FUNCTION "FRK_PersistDirty" : Void
{ S7_Optimized_Access := 'TRUE' }
VERSION : 0.1
VAR_INPUT
    Slot : Int;
END_VAR
VAR_TEMP
    Stamp : LDT;
    NativeResult : Int;
END_VAR
BEGIN
    IF #Slot < 1 OR #Slot > 20 THEN RETURN; END_IF;
    IF NOT "FRK_PersistConsumers".Rows[#Slot].Dirty THEN
        #NativeResult := RD_SYS_T(OUT => #Stamp);
        IF "FRK_PersistConsumers".Rows[#Slot].Ticket = 0 THEN "FRK_PersistConsumers".Rows[#Slot].PendingSince := #Stamp;
        ELSE "FRK_PersistConsumers".Rows[#Slot].NextSince := #Stamp; END_IF;
    END_IF;
    "FRK_PersistConsumers".Rows[#Slot].Dirty := TRUE;
END_FUNCTION
FUNCTION "FRK_PersistConfigSlot" : Int
{ S7_Optimized_Access := 'TRUE' }
VERSION : 0.1
VAR_INPUT
    Scope : String;
    ModelCode : String;
    Kind : DInt;
END_VAR
BEGIN
    #FRK_PersistConfigSlot := 0;
    IF #Scope = 'StationA' AND #ModelCode = '' AND #Kind = 1 THEN #FRK_PersistConfigSlot := 1; RETURN; END_IF;
    IF #Scope = 'StationA' AND #ModelCode = '' AND #Kind = 1 THEN #FRK_PersistConfigSlot := 1; RETURN; END_IF;
    IF #Scope = 'StationA' AND #ModelCode = '' AND #Kind = 1 THEN #FRK_PersistConfigSlot := 1; RETURN; END_IF;
    IF #Scope = 'StationA' AND #ModelCode = '' AND #Kind = 1 THEN #FRK_PersistConfigSlot := 1; RETURN; END_IF;
    IF #Scope = 'StationA' AND #ModelCode = '' AND #Kind = 1 THEN #FRK_PersistConfigSlot := 1; RETURN; END_IF;
    IF #Scope = 'StationA' AND #ModelCode = '' AND #Kind = 1 THEN #FRK_PersistConfigSlot := 1; RETURN; END_IF;
    IF #Scope = 'StationA' AND #ModelCode = '' AND #Kind = 1 THEN #FRK_PersistConfigSlot := 1; RETURN; END_IF;
    IF #Scope = 'StationA' AND #ModelCode = '' AND #Kind = 1 THEN #FRK_PersistConfigSlot := 1; RETURN; END_IF;
    IF #Scope = 'StationA.Satellite' AND #ModelCode = '' AND #Kind = 1 THEN #FRK_PersistConfigSlot := 1; RETURN; END_IF;
    IF #Scope = 'StationA.Satellite' AND #ModelCode = '' AND #Kind = 1 THEN #FRK_PersistConfigSlot := 1; RETURN; END_IF;
    IF #Scope = 'StationA.Satellite' AND #ModelCode = '' AND #Kind = 1 THEN #FRK_PersistConfigSlot := 1; RETURN; END_IF;
    IF #Scope = 'StationA.Satellite' AND #ModelCode = '' AND #Kind = 1 THEN #FRK_PersistConfigSlot := 1; RETURN; END_IF;
    IF #Scope = 'StationA.Satellite' AND #ModelCode = '' AND #Kind = 1 THEN #FRK_PersistConfigSlot := 1; RETURN; END_IF;
    IF #Scope = 'StationA.Satellite' AND #ModelCode = '' AND #Kind = 1 THEN #FRK_PersistConfigSlot := 1; RETURN; END_IF;
    IF #Scope = 'StationA.Satellite' AND #ModelCode = '' AND #Kind = 1 THEN #FRK_PersistConfigSlot := 1; RETURN; END_IF;
    IF #Scope = 'StationA.Satellite' AND #ModelCode = '' AND #Kind = 1 THEN #FRK_PersistConfigSlot := 1; RETURN; END_IF;
    IF #Scope = 'StationA.Satellite' AND #ModelCode = '' AND #Kind = 1 THEN #FRK_PersistConfigSlot := 1; RETURN; END_IF;
    IF #Scope = 'StationA.Satellite' AND #ModelCode = '' AND #Kind = 1 THEN #FRK_PersistConfigSlot := 1; RETURN; END_IF;
    IF #Scope = 'StationA.Satellite.Inner' AND #ModelCode = '' AND #Kind = 1 THEN #FRK_PersistConfigSlot := 1; RETURN; END_IF;
    IF #Scope = 'StationA.Satellite.Inner' AND #ModelCode = '' AND #Kind = 1 THEN #FRK_PersistConfigSlot := 1; RETURN; END_IF;
    IF #Scope = 'StationA.Satellite.Inner' AND #ModelCode = '' AND #Kind = 1 THEN #FRK_PersistConfigSlot := 1; RETURN; END_IF;
    IF #Scope = 'StationA.Satellite.Inner' AND #ModelCode = '' AND #Kind = 1 THEN #FRK_PersistConfigSlot := 1; RETURN; END_IF;
    IF #Scope = 'StationA.Satellite.Inner' AND #ModelCode = '' AND #Kind = 1 THEN #FRK_PersistConfigSlot := 1; RETURN; END_IF;
    IF #Scope = 'StationA.Satellite.Inner' AND #ModelCode = '' AND #Kind = 1 THEN #FRK_PersistConfigSlot := 1; RETURN; END_IF;
    IF #Scope = 'StationA.Satellite.Inner' AND #ModelCode = '' AND #Kind = 1 THEN #FRK_PersistConfigSlot := 1; RETURN; END_IF;
    IF #Scope = 'StationA.Satellite.Inner' AND #ModelCode = '' AND #Kind = 1 THEN #FRK_PersistConfigSlot := 1; RETURN; END_IF;
    IF #Scope = 'StationA.Satellite.Inner' AND #ModelCode = '' AND #Kind = 1 THEN #FRK_PersistConfigSlot := 1; RETURN; END_IF;
    IF #Scope = 'StationA.Satellite.Inner' AND #ModelCode = '' AND #Kind = 1 THEN #FRK_PersistConfigSlot := 1; RETURN; END_IF;
    IF #Scope = 'StationA' AND #ModelCode = 'MODEL_A' AND #Kind = 0 THEN #FRK_PersistConfigSlot := 2; RETURN; END_IF;
    IF #Scope = 'StationA' AND #ModelCode = 'MODEL_A' AND #Kind = 0 THEN #FRK_PersistConfigSlot := 2; RETURN; END_IF;
    IF #Scope = 'StationA' AND #ModelCode = 'MODEL_A' AND #Kind = 0 THEN #FRK_PersistConfigSlot := 2; RETURN; END_IF;
    IF #Scope = 'StationA' AND #ModelCode = 'MODEL_A' AND #Kind = 0 THEN #FRK_PersistConfigSlot := 2; RETURN; END_IF;
    IF #Scope = 'StationA.Cell' AND #ModelCode = 'MODEL_A' AND #Kind = 0 THEN #FRK_PersistConfigSlot := 2; RETURN; END_IF;
    IF #Scope = 'StationA.Cell' AND #ModelCode = 'MODEL_A' AND #Kind = 0 THEN #FRK_PersistConfigSlot := 2; RETURN; END_IF;
    IF #Scope = 'StationA.Cell.Clamp' AND #ModelCode = 'MODEL_A' AND #Kind = 0 THEN #FRK_PersistConfigSlot := 2; RETURN; END_IF;
    IF #Scope = 'StationA.Cell.Clamp' AND #ModelCode = 'MODEL_A' AND #Kind = 0 THEN #FRK_PersistConfigSlot := 2; RETURN; END_IF;
    IF #Scope = 'StationA.Cell.Gate' AND #ModelCode = 'MODEL_A' AND #Kind = 0 THEN #FRK_PersistConfigSlot := 2; RETURN; END_IF;
    IF #Scope = 'StationA.Cell.Gate' AND #ModelCode = 'MODEL_A' AND #Kind = 0 THEN #FRK_PersistConfigSlot := 2; RETURN; END_IF;
    IF #Scope = 'StationA.Satellite' AND #ModelCode = 'MODEL_A' AND #Kind = 0 THEN #FRK_PersistConfigSlot := 2; RETURN; END_IF;
    IF #Scope = 'StationA.Satellite' AND #ModelCode = 'MODEL_A' AND #Kind = 0 THEN #FRK_PersistConfigSlot := 2; RETURN; END_IF;
    IF #Scope = 'StationA.Satellite.Cell' AND #ModelCode = 'MODEL_A' AND #Kind = 0 THEN #FRK_PersistConfigSlot := 2; RETURN; END_IF;
    IF #Scope = 'StationA.Satellite.Cell' AND #ModelCode = 'MODEL_A' AND #Kind = 0 THEN #FRK_PersistConfigSlot := 2; RETURN; END_IF;
    IF #Scope = 'StationA.Satellite.Cell.Clamp' AND #ModelCode = 'MODEL_A' AND #Kind = 0 THEN #FRK_PersistConfigSlot := 2; RETURN; END_IF;
    IF #Scope = 'StationA.Satellite.Cell.Clamp' AND #ModelCode = 'MODEL_A' AND #Kind = 0 THEN #FRK_PersistConfigSlot := 2; RETURN; END_IF;
    IF #Scope = 'StationA.Satellite.Cell.Gate' AND #ModelCode = 'MODEL_A' AND #Kind = 0 THEN #FRK_PersistConfigSlot := 2; RETURN; END_IF;
    IF #Scope = 'StationA.Satellite.Cell.Gate' AND #ModelCode = 'MODEL_A' AND #Kind = 0 THEN #FRK_PersistConfigSlot := 2; RETURN; END_IF;
    IF #Scope = 'StationA.Satellite.Inner' AND #ModelCode = 'MODEL_A' AND #Kind = 0 THEN #FRK_PersistConfigSlot := 2; RETURN; END_IF;
    IF #Scope = 'StationA.Satellite.Inner' AND #ModelCode = 'MODEL_A' AND #Kind = 0 THEN #FRK_PersistConfigSlot := 2; RETURN; END_IF;
    IF #Scope = 'StationA.Satellite.Inner.Cell' AND #ModelCode = 'MODEL_A' AND #Kind = 0 THEN #FRK_PersistConfigSlot := 2; RETURN; END_IF;
    IF #Scope = 'StationA.Satellite.Inner.Cell' AND #ModelCode = 'MODEL_A' AND #Kind = 0 THEN #FRK_PersistConfigSlot := 2; RETURN; END_IF;
    IF #Scope = 'StationA.Satellite.Inner.Cell.Clamp' AND #ModelCode = 'MODEL_A' AND #Kind = 0 THEN #FRK_PersistConfigSlot := 2; RETURN; END_IF;
    IF #Scope = 'StationA.Satellite.Inner.Cell.Clamp' AND #ModelCode = 'MODEL_A' AND #Kind = 0 THEN #FRK_PersistConfigSlot := 2; RETURN; END_IF;
    IF #Scope = 'StationA.Satellite.Inner.Cell.Gate' AND #ModelCode = 'MODEL_A' AND #Kind = 0 THEN #FRK_PersistConfigSlot := 2; RETURN; END_IF;
    IF #Scope = 'StationA.Satellite.Inner.Cell.Gate' AND #ModelCode = 'MODEL_A' AND #Kind = 0 THEN #FRK_PersistConfigSlot := 2; RETURN; END_IF;
    IF #Scope = 'StationA' AND #ModelCode = 'MODEL_B' AND #Kind = 0 THEN #FRK_PersistConfigSlot := 3; RETURN; END_IF;
    IF #Scope = 'StationA' AND #ModelCode = 'MODEL_B' AND #Kind = 0 THEN #FRK_PersistConfigSlot := 3; RETURN; END_IF;
    IF #Scope = 'StationA' AND #ModelCode = 'MODEL_B' AND #Kind = 0 THEN #FRK_PersistConfigSlot := 3; RETURN; END_IF;
    IF #Scope = 'StationA' AND #ModelCode = 'MODEL_B' AND #Kind = 0 THEN #FRK_PersistConfigSlot := 3; RETURN; END_IF;
    IF #Scope = 'StationA.Cell' AND #ModelCode = 'MODEL_B' AND #Kind = 0 THEN #FRK_PersistConfigSlot := 3; RETURN; END_IF;
    IF #Scope = 'StationA.Cell' AND #ModelCode = 'MODEL_B' AND #Kind = 0 THEN #FRK_PersistConfigSlot := 3; RETURN; END_IF;
    IF #Scope = 'StationA.Cell.Clamp' AND #ModelCode = 'MODEL_B' AND #Kind = 0 THEN #FRK_PersistConfigSlot := 3; RETURN; END_IF;
    IF #Scope = 'StationA.Cell.Clamp' AND #ModelCode = 'MODEL_B' AND #Kind = 0 THEN #FRK_PersistConfigSlot := 3; RETURN; END_IF;
    IF #Scope = 'StationA.Cell.Gate' AND #ModelCode = 'MODEL_B' AND #Kind = 0 THEN #FRK_PersistConfigSlot := 3; RETURN; END_IF;
    IF #Scope = 'StationA.Cell.Gate' AND #ModelCode = 'MODEL_B' AND #Kind = 0 THEN #FRK_PersistConfigSlot := 3; RETURN; END_IF;
    IF #Scope = 'StationA.Satellite' AND #ModelCode = 'MODEL_B' AND #Kind = 0 THEN #FRK_PersistConfigSlot := 3; RETURN; END_IF;
    IF #Scope = 'StationA.Satellite' AND #ModelCode = 'MODEL_B' AND #Kind = 0 THEN #FRK_PersistConfigSlot := 3; RETURN; END_IF;
    IF #Scope = 'StationA.Satellite.Cell' AND #ModelCode = 'MODEL_B' AND #Kind = 0 THEN #FRK_PersistConfigSlot := 3; RETURN; END_IF;
    IF #Scope = 'StationA.Satellite.Cell' AND #ModelCode = 'MODEL_B' AND #Kind = 0 THEN #FRK_PersistConfigSlot := 3; RETURN; END_IF;
    IF #Scope = 'StationA.Satellite.Cell.Clamp' AND #ModelCode = 'MODEL_B' AND #Kind = 0 THEN #FRK_PersistConfigSlot := 3; RETURN; END_IF;
    IF #Scope = 'StationA.Satellite.Cell.Clamp' AND #ModelCode = 'MODEL_B' AND #Kind = 0 THEN #FRK_PersistConfigSlot := 3; RETURN; END_IF;
    IF #Scope = 'StationA.Satellite.Cell.Gate' AND #ModelCode = 'MODEL_B' AND #Kind = 0 THEN #FRK_PersistConfigSlot := 3; RETURN; END_IF;
    IF #Scope = 'StationA.Satellite.Cell.Gate' AND #ModelCode = 'MODEL_B' AND #Kind = 0 THEN #FRK_PersistConfigSlot := 3; RETURN; END_IF;
    IF #Scope = 'StationA.Satellite.Inner' AND #ModelCode = 'MODEL_B' AND #Kind = 0 THEN #FRK_PersistConfigSlot := 3; RETURN; END_IF;
    IF #Scope = 'StationA.Satellite.Inner' AND #ModelCode = 'MODEL_B' AND #Kind = 0 THEN #FRK_PersistConfigSlot := 3; RETURN; END_IF;
    IF #Scope = 'StationA.Satellite.Inner.Cell' AND #ModelCode = 'MODEL_B' AND #Kind = 0 THEN #FRK_PersistConfigSlot := 3; RETURN; END_IF;
    IF #Scope = 'StationA.Satellite.Inner.Cell' AND #ModelCode = 'MODEL_B' AND #Kind = 0 THEN #FRK_PersistConfigSlot := 3; RETURN; END_IF;
    IF #Scope = 'StationA.Satellite.Inner.Cell.Clamp' AND #ModelCode = 'MODEL_B' AND #Kind = 0 THEN #FRK_PersistConfigSlot := 3; RETURN; END_IF;
    IF #Scope = 'StationA.Satellite.Inner.Cell.Clamp' AND #ModelCode = 'MODEL_B' AND #Kind = 0 THEN #FRK_PersistConfigSlot := 3; RETURN; END_IF;
    IF #Scope = 'StationA.Satellite.Inner.Cell.Gate' AND #ModelCode = 'MODEL_B' AND #Kind = 0 THEN #FRK_PersistConfigSlot := 3; RETURN; END_IF;
    IF #Scope = 'StationA.Satellite.Inner.Cell.Gate' AND #ModelCode = 'MODEL_B' AND #Kind = 0 THEN #FRK_PersistConfigSlot := 3; RETURN; END_IF;
    IF #Scope = 'StationB' AND #ModelCode = '' AND #Kind = 1 THEN #FRK_PersistConfigSlot := 9; RETURN; END_IF;
    IF #Scope = 'StationB' AND #ModelCode = '' AND #Kind = 1 THEN #FRK_PersistConfigSlot := 9; RETURN; END_IF;
    IF #Scope = 'StationB' AND #ModelCode = '' AND #Kind = 1 THEN #FRK_PersistConfigSlot := 9; RETURN; END_IF;
    IF #Scope = 'StationB' AND #ModelCode = '' AND #Kind = 1 THEN #FRK_PersistConfigSlot := 9; RETURN; END_IF;
    IF #Scope = 'StationB' AND #ModelCode = '' AND #Kind = 1 THEN #FRK_PersistConfigSlot := 9; RETURN; END_IF;
    IF #Scope = 'StationB' AND #ModelCode = '' AND #Kind = 1 THEN #FRK_PersistConfigSlot := 9; RETURN; END_IF;
    IF #Scope = 'StationB' AND #ModelCode = '' AND #Kind = 1 THEN #FRK_PersistConfigSlot := 9; RETURN; END_IF;
    IF #Scope = 'StationB' AND #ModelCode = '' AND #Kind = 1 THEN #FRK_PersistConfigSlot := 9; RETURN; END_IF;
    IF #Scope = 'StationB.Satellite' AND #ModelCode = '' AND #Kind = 1 THEN #FRK_PersistConfigSlot := 9; RETURN; END_IF;
    IF #Scope = 'StationB.Satellite' AND #ModelCode = '' AND #Kind = 1 THEN #FRK_PersistConfigSlot := 9; RETURN; END_IF;
    IF #Scope = 'StationB.Satellite' AND #ModelCode = '' AND #Kind = 1 THEN #FRK_PersistConfigSlot := 9; RETURN; END_IF;
    IF #Scope = 'StationB.Satellite' AND #ModelCode = '' AND #Kind = 1 THEN #FRK_PersistConfigSlot := 9; RETURN; END_IF;
    IF #Scope = 'StationB.Satellite' AND #ModelCode = '' AND #Kind = 1 THEN #FRK_PersistConfigSlot := 9; RETURN; END_IF;
    IF #Scope = 'StationB.Satellite' AND #ModelCode = '' AND #Kind = 1 THEN #FRK_PersistConfigSlot := 9; RETURN; END_IF;
    IF #Scope = 'StationB.Satellite' AND #ModelCode = '' AND #Kind = 1 THEN #FRK_PersistConfigSlot := 9; RETURN; END_IF;
    IF #Scope = 'StationB.Satellite' AND #ModelCode = '' AND #Kind = 1 THEN #FRK_PersistConfigSlot := 9; RETURN; END_IF;
    IF #Scope = 'StationB.Satellite' AND #ModelCode = '' AND #Kind = 1 THEN #FRK_PersistConfigSlot := 9; RETURN; END_IF;
    IF #Scope = 'StationB.Satellite' AND #ModelCode = '' AND #Kind = 1 THEN #FRK_PersistConfigSlot := 9; RETURN; END_IF;
    IF #Scope = 'StationB.Satellite.Inner' AND #ModelCode = '' AND #Kind = 1 THEN #FRK_PersistConfigSlot := 9; RETURN; END_IF;
    IF #Scope = 'StationB.Satellite.Inner' AND #ModelCode = '' AND #Kind = 1 THEN #FRK_PersistConfigSlot := 9; RETURN; END_IF;
    IF #Scope = 'StationB.Satellite.Inner' AND #ModelCode = '' AND #Kind = 1 THEN #FRK_PersistConfigSlot := 9; RETURN; END_IF;
    IF #Scope = 'StationB.Satellite.Inner' AND #ModelCode = '' AND #Kind = 1 THEN #FRK_PersistConfigSlot := 9; RETURN; END_IF;
    IF #Scope = 'StationB.Satellite.Inner' AND #ModelCode = '' AND #Kind = 1 THEN #FRK_PersistConfigSlot := 9; RETURN; END_IF;
    IF #Scope = 'StationB.Satellite.Inner' AND #ModelCode = '' AND #Kind = 1 THEN #FRK_PersistConfigSlot := 9; RETURN; END_IF;
    IF #Scope = 'StationB.Satellite.Inner' AND #ModelCode = '' AND #Kind = 1 THEN #FRK_PersistConfigSlot := 9; RETURN; END_IF;
    IF #Scope = 'StationB.Satellite.Inner' AND #ModelCode = '' AND #Kind = 1 THEN #FRK_PersistConfigSlot := 9; RETURN; END_IF;
    IF #Scope = 'StationB.Satellite.Inner' AND #ModelCode = '' AND #Kind = 1 THEN #FRK_PersistConfigSlot := 9; RETURN; END_IF;
    IF #Scope = 'StationB.Satellite.Inner' AND #ModelCode = '' AND #Kind = 1 THEN #FRK_PersistConfigSlot := 9; RETURN; END_IF;
    IF #Scope = 'StationB' AND #ModelCode = 'MODEL_A' AND #Kind = 0 THEN #FRK_PersistConfigSlot := 10; RETURN; END_IF;
    IF #Scope = 'StationB' AND #ModelCode = 'MODEL_A' AND #Kind = 0 THEN #FRK_PersistConfigSlot := 10; RETURN; END_IF;
    IF #Scope = 'StationB' AND #ModelCode = 'MODEL_A' AND #Kind = 0 THEN #FRK_PersistConfigSlot := 10; RETURN; END_IF;
    IF #Scope = 'StationB' AND #ModelCode = 'MODEL_A' AND #Kind = 0 THEN #FRK_PersistConfigSlot := 10; RETURN; END_IF;
    IF #Scope = 'StationB.Cell' AND #ModelCode = 'MODEL_A' AND #Kind = 0 THEN #FRK_PersistConfigSlot := 10; RETURN; END_IF;
    IF #Scope = 'StationB.Cell' AND #ModelCode = 'MODEL_A' AND #Kind = 0 THEN #FRK_PersistConfigSlot := 10; RETURN; END_IF;
    IF #Scope = 'StationB.Cell.Clamp' AND #ModelCode = 'MODEL_A' AND #Kind = 0 THEN #FRK_PersistConfigSlot := 10; RETURN; END_IF;
    IF #Scope = 'StationB.Cell.Clamp' AND #ModelCode = 'MODEL_A' AND #Kind = 0 THEN #FRK_PersistConfigSlot := 10; RETURN; END_IF;
    IF #Scope = 'StationB.Cell.Gate' AND #ModelCode = 'MODEL_A' AND #Kind = 0 THEN #FRK_PersistConfigSlot := 10; RETURN; END_IF;
    IF #Scope = 'StationB.Cell.Gate' AND #ModelCode = 'MODEL_A' AND #Kind = 0 THEN #FRK_PersistConfigSlot := 10; RETURN; END_IF;
    IF #Scope = 'StationB.Satellite' AND #ModelCode = 'MODEL_A' AND #Kind = 0 THEN #FRK_PersistConfigSlot := 10; RETURN; END_IF;
    IF #Scope = 'StationB.Satellite' AND #ModelCode = 'MODEL_A' AND #Kind = 0 THEN #FRK_PersistConfigSlot := 10; RETURN; END_IF;
    IF #Scope = 'StationB.Satellite.Cell' AND #ModelCode = 'MODEL_A' AND #Kind = 0 THEN #FRK_PersistConfigSlot := 10; RETURN; END_IF;
    IF #Scope = 'StationB.Satellite.Cell' AND #ModelCode = 'MODEL_A' AND #Kind = 0 THEN #FRK_PersistConfigSlot := 10; RETURN; END_IF;
    IF #Scope = 'StationB.Satellite.Cell.Clamp' AND #ModelCode = 'MODEL_A' AND #Kind = 0 THEN #FRK_PersistConfigSlot := 10; RETURN; END_IF;
    IF #Scope = 'StationB.Satellite.Cell.Clamp' AND #ModelCode = 'MODEL_A' AND #Kind = 0 THEN #FRK_PersistConfigSlot := 10; RETURN; END_IF;
    IF #Scope = 'StationB.Satellite.Cell.Gate' AND #ModelCode = 'MODEL_A' AND #Kind = 0 THEN #FRK_PersistConfigSlot := 10; RETURN; END_IF;
    IF #Scope = 'StationB.Satellite.Cell.Gate' AND #ModelCode = 'MODEL_A' AND #Kind = 0 THEN #FRK_PersistConfigSlot := 10; RETURN; END_IF;
    IF #Scope = 'StationB.Satellite.Inner' AND #ModelCode = 'MODEL_A' AND #Kind = 0 THEN #FRK_PersistConfigSlot := 10; RETURN; END_IF;
    IF #Scope = 'StationB.Satellite.Inner' AND #ModelCode = 'MODEL_A' AND #Kind = 0 THEN #FRK_PersistConfigSlot := 10; RETURN; END_IF;
    IF #Scope = 'StationB.Satellite.Inner.Cell' AND #ModelCode = 'MODEL_A' AND #Kind = 0 THEN #FRK_PersistConfigSlot := 10; RETURN; END_IF;
    IF #Scope = 'StationB.Satellite.Inner.Cell' AND #ModelCode = 'MODEL_A' AND #Kind = 0 THEN #FRK_PersistConfigSlot := 10; RETURN; END_IF;
    IF #Scope = 'StationB.Satellite.Inner.Cell.Clamp' AND #ModelCode = 'MODEL_A' AND #Kind = 0 THEN #FRK_PersistConfigSlot := 10; RETURN; END_IF;
    IF #Scope = 'StationB.Satellite.Inner.Cell.Clamp' AND #ModelCode = 'MODEL_A' AND #Kind = 0 THEN #FRK_PersistConfigSlot := 10; RETURN; END_IF;
    IF #Scope = 'StationB.Satellite.Inner.Cell.Gate' AND #ModelCode = 'MODEL_A' AND #Kind = 0 THEN #FRK_PersistConfigSlot := 10; RETURN; END_IF;
    IF #Scope = 'StationB.Satellite.Inner.Cell.Gate' AND #ModelCode = 'MODEL_A' AND #Kind = 0 THEN #FRK_PersistConfigSlot := 10; RETURN; END_IF;
    IF #Scope = 'StationB' AND #ModelCode = 'MODEL_B' AND #Kind = 0 THEN #FRK_PersistConfigSlot := 11; RETURN; END_IF;
    IF #Scope = 'StationB' AND #ModelCode = 'MODEL_B' AND #Kind = 0 THEN #FRK_PersistConfigSlot := 11; RETURN; END_IF;
    IF #Scope = 'StationB' AND #ModelCode = 'MODEL_B' AND #Kind = 0 THEN #FRK_PersistConfigSlot := 11; RETURN; END_IF;
    IF #Scope = 'StationB' AND #ModelCode = 'MODEL_B' AND #Kind = 0 THEN #FRK_PersistConfigSlot := 11; RETURN; END_IF;
    IF #Scope = 'StationB.Cell' AND #ModelCode = 'MODEL_B' AND #Kind = 0 THEN #FRK_PersistConfigSlot := 11; RETURN; END_IF;
    IF #Scope = 'StationB.Cell' AND #ModelCode = 'MODEL_B' AND #Kind = 0 THEN #FRK_PersistConfigSlot := 11; RETURN; END_IF;
    IF #Scope = 'StationB.Cell.Clamp' AND #ModelCode = 'MODEL_B' AND #Kind = 0 THEN #FRK_PersistConfigSlot := 11; RETURN; END_IF;
    IF #Scope = 'StationB.Cell.Clamp' AND #ModelCode = 'MODEL_B' AND #Kind = 0 THEN #FRK_PersistConfigSlot := 11; RETURN; END_IF;
    IF #Scope = 'StationB.Cell.Gate' AND #ModelCode = 'MODEL_B' AND #Kind = 0 THEN #FRK_PersistConfigSlot := 11; RETURN; END_IF;
    IF #Scope = 'StationB.Cell.Gate' AND #ModelCode = 'MODEL_B' AND #Kind = 0 THEN #FRK_PersistConfigSlot := 11; RETURN; END_IF;
    IF #Scope = 'StationB.Satellite' AND #ModelCode = 'MODEL_B' AND #Kind = 0 THEN #FRK_PersistConfigSlot := 11; RETURN; END_IF;
    IF #Scope = 'StationB.Satellite' AND #ModelCode = 'MODEL_B' AND #Kind = 0 THEN #FRK_PersistConfigSlot := 11; RETURN; END_IF;
    IF #Scope = 'StationB.Satellite.Cell' AND #ModelCode = 'MODEL_B' AND #Kind = 0 THEN #FRK_PersistConfigSlot := 11; RETURN; END_IF;
    IF #Scope = 'StationB.Satellite.Cell' AND #ModelCode = 'MODEL_B' AND #Kind = 0 THEN #FRK_PersistConfigSlot := 11; RETURN; END_IF;
    IF #Scope = 'StationB.Satellite.Cell.Clamp' AND #ModelCode = 'MODEL_B' AND #Kind = 0 THEN #FRK_PersistConfigSlot := 11; RETURN; END_IF;
    IF #Scope = 'StationB.Satellite.Cell.Clamp' AND #ModelCode = 'MODEL_B' AND #Kind = 0 THEN #FRK_PersistConfigSlot := 11; RETURN; END_IF;
    IF #Scope = 'StationB.Satellite.Cell.Gate' AND #ModelCode = 'MODEL_B' AND #Kind = 0 THEN #FRK_PersistConfigSlot := 11; RETURN; END_IF;
    IF #Scope = 'StationB.Satellite.Cell.Gate' AND #ModelCode = 'MODEL_B' AND #Kind = 0 THEN #FRK_PersistConfigSlot := 11; RETURN; END_IF;
    IF #Scope = 'StationB.Satellite.Inner' AND #ModelCode = 'MODEL_B' AND #Kind = 0 THEN #FRK_PersistConfigSlot := 11; RETURN; END_IF;
    IF #Scope = 'StationB.Satellite.Inner' AND #ModelCode = 'MODEL_B' AND #Kind = 0 THEN #FRK_PersistConfigSlot := 11; RETURN; END_IF;
    IF #Scope = 'StationB.Satellite.Inner.Cell' AND #ModelCode = 'MODEL_B' AND #Kind = 0 THEN #FRK_PersistConfigSlot := 11; RETURN; END_IF;
    IF #Scope = 'StationB.Satellite.Inner.Cell' AND #ModelCode = 'MODEL_B' AND #Kind = 0 THEN #FRK_PersistConfigSlot := 11; RETURN; END_IF;
    IF #Scope = 'StationB.Satellite.Inner.Cell.Clamp' AND #ModelCode = 'MODEL_B' AND #Kind = 0 THEN #FRK_PersistConfigSlot := 11; RETURN; END_IF;
    IF #Scope = 'StationB.Satellite.Inner.Cell.Clamp' AND #ModelCode = 'MODEL_B' AND #Kind = 0 THEN #FRK_PersistConfigSlot := 11; RETURN; END_IF;
    IF #Scope = 'StationB.Satellite.Inner.Cell.Gate' AND #ModelCode = 'MODEL_B' AND #Kind = 0 THEN #FRK_PersistConfigSlot := 11; RETURN; END_IF;
    IF #Scope = 'StationB.Satellite.Inner.Cell.Gate' AND #ModelCode = 'MODEL_B' AND #Kind = 0 THEN #FRK_PersistConfigSlot := 11; RETURN; END_IF;
END_FUNCTION
FUNCTION "FRK_PersistUsersDirty" : Void
{ S7_Optimized_Access := 'TRUE' }
VERSION : 0.1
BEGIN
    "FRK_PersistDirty"(Slot := 17);
END_FUNCTION
FUNCTION "FRK_PersistPolicyDirty" : Void
{ S7_Optimized_Access := 'TRUE' }
VERSION : 0.1
VAR_INPUT
    RootIndex : Int;
END_VAR
BEGIN
    IF #RootIndex = 1 THEN "FRK_PersistDirty"(Slot := 4); END_IF;
    IF #RootIndex = 2 THEN "FRK_PersistDirty"(Slot := 12); END_IF;
END_FUNCTION
FUNCTION "FRK_PersistSetDirty" : Void
{ S7_Optimized_Access := 'TRUE' }
VERSION : 0.1
VAR_INPUT
    RootIndex : Int;
    Ordinal : Int;
END_VAR
BEGIN
    IF #RootIndex = 1 AND #Ordinal = 1 THEN "FRK_PersistDirty"(Slot := 5); END_IF;
    IF #RootIndex = 1 AND #Ordinal = 2 THEN "FRK_PersistDirty"(Slot := 6); END_IF;
    IF #RootIndex = 1 AND #Ordinal = 3 THEN "FRK_PersistDirty"(Slot := 7); END_IF;
    IF #RootIndex = 1 AND #Ordinal = 4 THEN "FRK_PersistDirty"(Slot := 8); END_IF;
    IF #RootIndex = 2 AND #Ordinal = 1 THEN "FRK_PersistDirty"(Slot := 13); END_IF;
    IF #RootIndex = 2 AND #Ordinal = 2 THEN "FRK_PersistDirty"(Slot := 14); END_IF;
    IF #RootIndex = 2 AND #Ordinal = 3 THEN "FRK_PersistDirty"(Slot := 15); END_IF;
    IF #RootIndex = 2 AND #Ordinal = 4 THEN "FRK_PersistDirty"(Slot := 16); END_IF;
END_FUNCTION
FUNCTION "FRK_PersistModelDirty" : Void
{ S7_Optimized_Access := 'TRUE' }
VERSION : 0.1
VAR_INPUT
    RootIndex : Int;
END_VAR
BEGIN
    IF #RootIndex = 1 THEN "FRK_PersistDirty"(Slot := 1); END_IF;
    IF #RootIndex = 2 THEN "FRK_PersistDirty"(Slot := 9); END_IF;
END_FUNCTION
FUNCTION "FRK_PersistClassesDirty" : Void
{ S7_Optimized_Access := 'TRUE' }
VERSION : 0.1
VAR_INPUT
    RootIndex : Int;
END_VAR
BEGIN
    IF #RootIndex = 1 THEN "FRK_PersistDirty"(Slot := 19); END_IF;
    IF #RootIndex = 2 THEN "FRK_PersistDirty"(Slot := 20); END_IF;
END_FUNCTION
FUNCTION "FRK_PersistVirginConfig" : Bool
{ S7_Optimized_Access := 'TRUE' }
VERSION : 0.1
VAR_INPUT
    Scope : String;
    ModelCode : String;
    Kind : DInt;
END_VAR
VAR_TEMP
    Slot : Int;
END_VAR
BEGIN
    #FRK_PersistVirginConfig := FALSE;
    #Slot := "FRK_PersistConfigSlot"(Scope := #Scope, ModelCode := #ModelCode, Kind := #Kind);
    IF #Slot > 0 THEN #FRK_PersistVirginConfig := "FRK_PersistConsumers".Rows[#Slot].Virgin; END_IF;
END_FUNCTION
FUNCTION "FRK_PersistLineTick" : Void
{ S7_Optimized_Access := 'TRUE' }
VERSION : 0.1
BEGIN
    IF "FRK_PersistConsumers".Ready AND "FRK_Line".Data.Dirty THEN
        "FRK_PersistDirty"(Slot := 18);
        "FRK_Line".Data.Dirty := FALSE;
    END_IF;
END_FUNCTION
